TYPE "FRK_Profiler_PressDemoUnit"
VERSION : 0.1
   STRUCT
      "LastCycle" : "FRK_CycleProfile_PressDemoUnit";
      "StepStats" : Array[1..23] of "ST_TimingRow";
      "StatsTruncated" : Bool;
      "LastCycleTime" : Time;
      "MinCycleTime" : Time;
      "History" : Array[1..60] of "ST_CycleSummary";
      "HistoryHead" : Int;
   END_STRUCT;
END_TYPE
